# EPICS substitutions: asynPortDriverETH32/Db/ETH32Motors.substitutions
# Expanded at build time into ETH32Motors.db (one set of records per motor).
# P, R, PORT and TIMEOUT are given when the IOC loads ETH32Motors.db.
file "ETH32Motor.template"
{
pattern
{ N,  ADDR }
{ 1,  0    }
{ 2,  1    }
{ 3,  2    }
{ 4,  3    }
{ 5,  4    }
{ 6,  5    }
{ 7,  6    }
{ 8,  7    }
}
